// LS Electric XG5000 project: 555
// PLC LSPLC

PROGRAM E2E_PICKNPLACE (task: 스캔 프로그램)

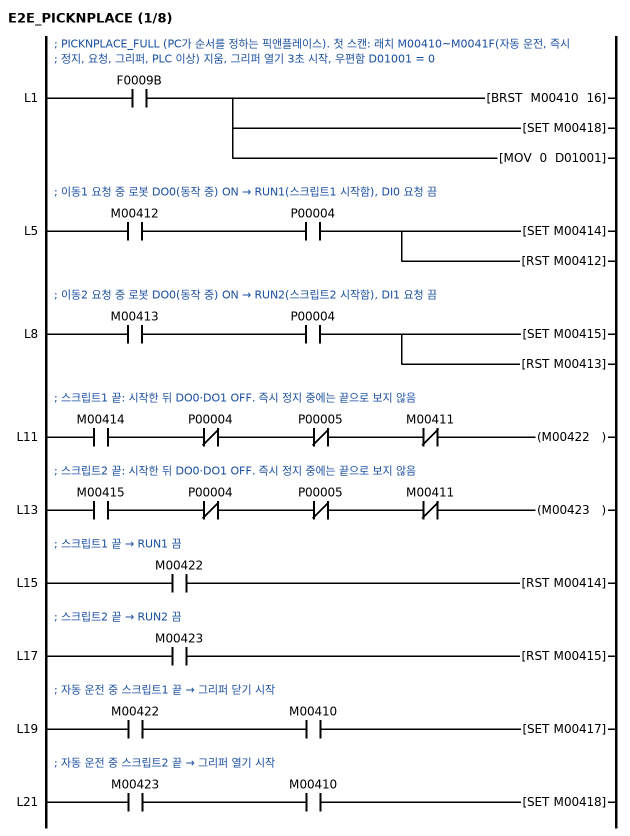
// PICKNPLACE_FULL (PC가 순서를 정하는 픽앤플레이스). 첫 스캔: 래치 M00410~M0041F(자동 운전, 즉시 정지, 요청, 그리퍼, PLC 이상) 지움, 그리퍼 열기 3초 시작, 우편함 D01001 = 0
; L1
LOAD      F0009B
BRST      M00410 16
SET       M00418
MOV       0 D01001
// 이동1 요청 중 로봇 DO0(동작 중) ON → RUN1(스크립트1 시작함), DI0 요청 끔
; L5
LOAD      M00412
AND       P00004
SET       M00414
RST       M00412
// 이동2 요청 중 로봇 DO0(동작 중) ON → RUN2(스크립트2 시작함), DI1 요청 끔
; L8
LOAD      M00413
AND       P00004
SET       M00415
RST       M00413
// 스크립트1 끝: 시작한 뒤 DO0·DO1 OFF. 즉시 정지 중에는 끝으로 보지 않음
; L11
LOAD      M00414
AND NOT   P00004
AND NOT   P00005
AND NOT   M00411
OUT       M00422
// 스크립트2 끝: 시작한 뒤 DO0·DO1 OFF. 즉시 정지 중에는 끝으로 보지 않음
; L13
LOAD      M00415
AND NOT   P00004
AND NOT   P00005
AND NOT   M00411
OUT       M00423
// 스크립트1 끝 → RUN1 끔
; L15
LOAD      M00422
RST       M00414
// 스크립트2 끝 → RUN2 끔
; L17
LOAD      M00423
RST       M00415
// 자동 운전 중 스크립트1 끝 → 그리퍼 닫기 시작
; L19
LOAD      M00422
AND       M00410
SET       M00417
// 자동 운전 중 스크립트2 끝 → 그리퍼 열기 시작
; L21
LOAD      M00423
AND       M00410
SET       M00418

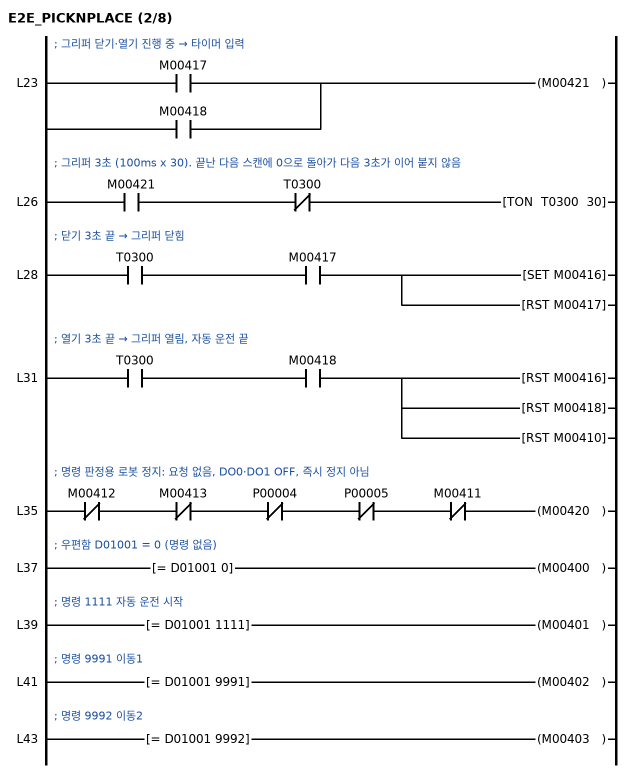
// 그리퍼 닫기·열기 진행 중 → 타이머 입력
; L23
LOAD      M00417
OR        M00418
OUT       M00421
// 그리퍼 3초 (100ms x 30). 끝난 다음 스캔에 0으로 돌아가 다음 3초가 이어 붙지 않음
; L26
LOAD      M00421
AND NOT   T0300
TON       T0300 30
// 닫기 3초 끝 → 그리퍼 닫힘
; L28
LOAD      T0300
AND       M00417
SET       M00416
RST       M00417
// 열기 3초 끝 → 그리퍼 열림, 자동 운전 끝
; L31
LOAD      T0300
AND       M00418
RST       M00416
RST       M00418
RST       M00410
// 명령 판정용 로봇 정지: 요청 없음, DO0·DO1 OFF, 즉시 정지 아님
; L35
LOAD NOT  M00412
AND NOT   M00413
AND NOT   P00004
AND NOT   P00005
AND NOT   M00411
OUT       M00420
// 우편함 D01001 = 0 (명령 없음)
; L37
LOAD=     D01001 0
OUT       M00400
// 명령 1111 자동 운전 시작
; L39
LOAD=     D01001 1111
OUT       M00401
// 명령 9991 이동1
; L41
LOAD=     D01001 9991
OUT       M00402
// 명령 9992 이동2
; L43
LOAD=     D01001 9992
OUT       M00403

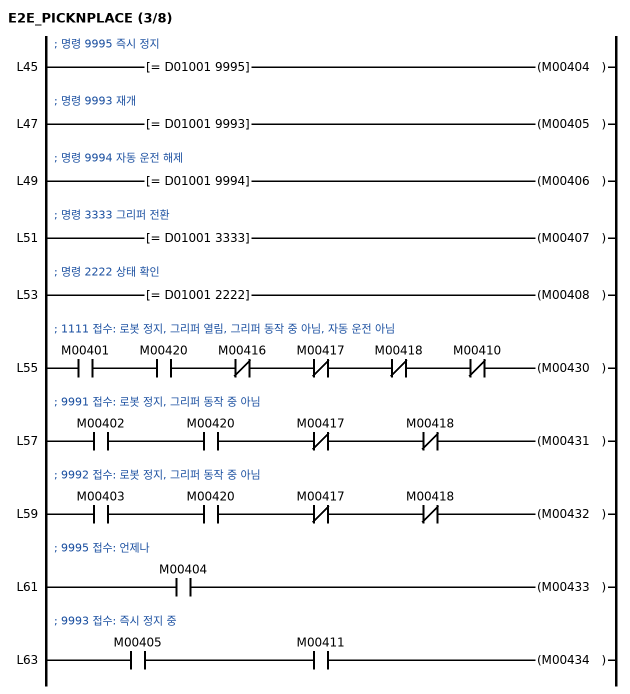
// 명령 9995 즉시 정지
; L45
LOAD=     D01001 9995
OUT       M00404
// 명령 9993 재개
; L47
LOAD=     D01001 9993
OUT       M00405
// 명령 9994 자동 운전 해제
; L49
LOAD=     D01001 9994
OUT       M00406
// 명령 3333 그리퍼 전환
; L51
LOAD=     D01001 3333
OUT       M00407
// 명령 2222 상태 확인
; L53
LOAD=     D01001 2222
OUT       M00408
// 1111 접수: 로봇 정지, 그리퍼 열림, 그리퍼 동작 중 아님, 자동 운전 아님
; L55
LOAD      M00401
AND       M00420
AND NOT   M00416
AND NOT   M00417
AND NOT   M00418
AND NOT   M00410
OUT       M00430
// 9991 접수: 로봇 정지, 그리퍼 동작 중 아님
; L57
LOAD      M00402
AND       M00420
AND NOT   M00417
AND NOT   M00418
OUT       M00431
// 9992 접수: 로봇 정지, 그리퍼 동작 중 아님
; L59
LOAD      M00403
AND       M00420
AND NOT   M00417
AND NOT   M00418
OUT       M00432
// 9995 접수: 언제나
; L61
LOAD      M00404
OUT       M00433
// 9993 접수: 즉시 정지 중
; L63
LOAD      M00405
AND       M00411
OUT       M00434

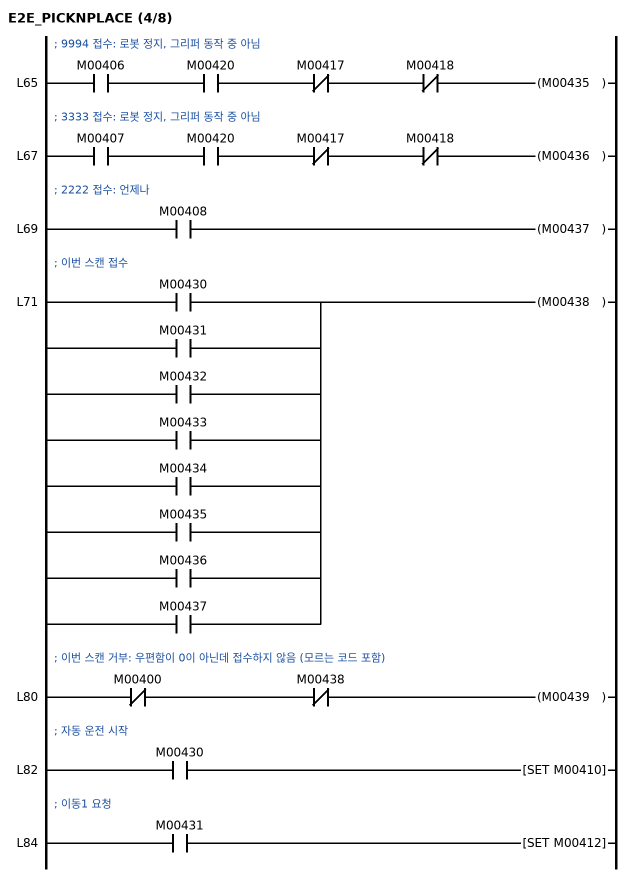
// 9994 접수: 로봇 정지, 그리퍼 동작 중 아님
; L65
LOAD      M00406
AND       M00420
AND NOT   M00417
AND NOT   M00418
OUT       M00435
// 3333 접수: 로봇 정지, 그리퍼 동작 중 아님
; L67
LOAD      M00407
AND       M00420
AND NOT   M00417
AND NOT   M00418
OUT       M00436
// 2222 접수: 언제나
; L69
LOAD      M00408
OUT       M00437
// 이번 스캔 접수
; L71
LOAD      M00430
OR        M00431
OR        M00432
OR        M00433
OR        M00434
OR        M00435
OR        M00436
OR        M00437
OUT       M00438
// 이번 스캔 거부: 우편함이 0이 아닌데 접수하지 않음 (모르는 코드 포함)
; L80
LOAD NOT  M00400
AND NOT   M00438
OUT       M00439
// 자동 운전 시작
; L82
LOAD      M00430
SET       M00410
// 이동1 요청
; L84
LOAD      M00431
SET       M00412

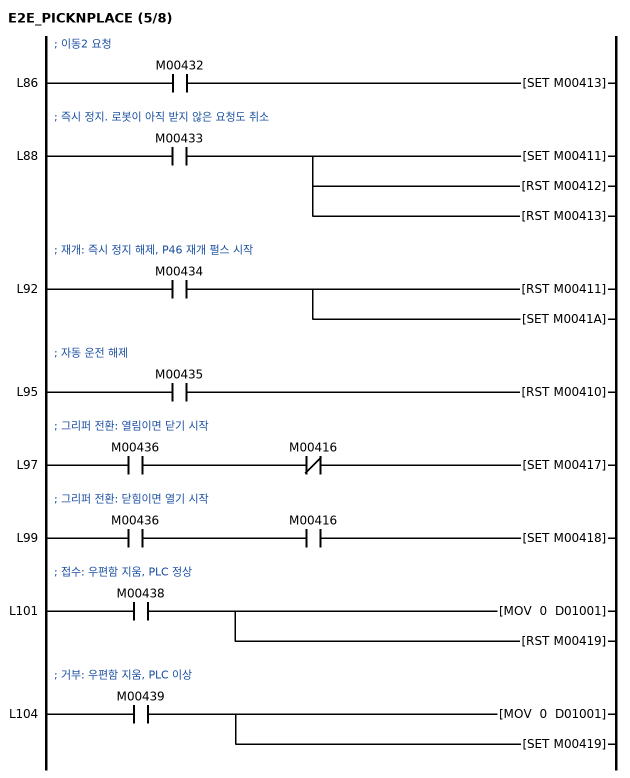
// 이동2 요청
; L86
LOAD      M00432
SET       M00413
// 즉시 정지. 로봇이 아직 받지 않은 요청도 취소
; L88
LOAD      M00433
SET       M00411
RST       M00412
RST       M00413
// 재개: 즉시 정지 해제, P46 재개 펄스 시작
; L92
LOAD      M00434
RST       M00411
SET       M0041A
// 자동 운전 해제
; L95
LOAD      M00435
RST       M00410
// 그리퍼 전환: 열림이면 닫기 시작
; L97
LOAD      M00436
AND NOT   M00416
SET       M00417
// 그리퍼 전환: 닫힘이면 열기 시작
; L99
LOAD      M00436
AND       M00416
SET       M00418
// 접수: 우편함 지움, PLC 정상
; L101
LOAD      M00438
MOV       0 D01001
RST       M00419
// 거부: 우편함 지움, PLC 이상
; L104
LOAD      M00439
MOV       0 D01001
SET       M00419

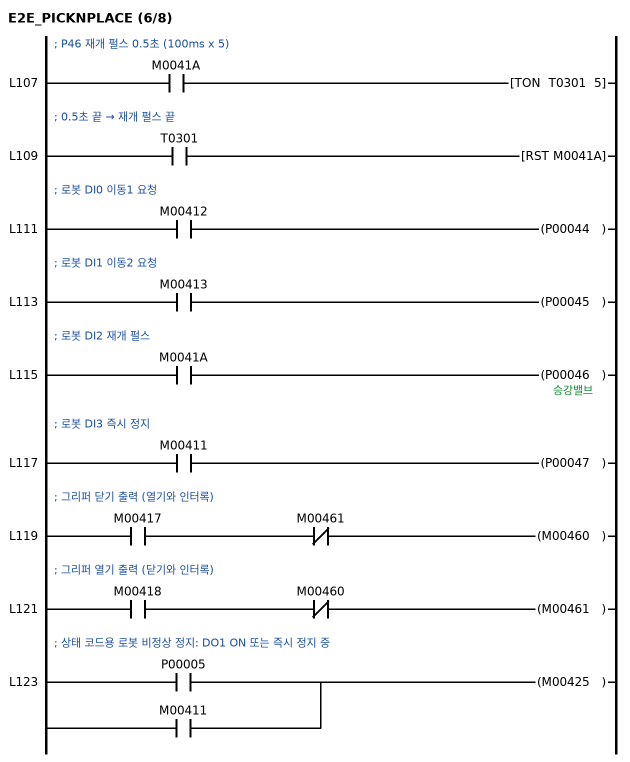
// P46 재개 펄스 0.5초 (100ms x 5)
; L107
LOAD      M0041A
TON       T0301 5
// 0.5초 끝 → 재개 펄스 끝
; L109
LOAD      T0301
RST       M0041A
// 로봇 DI0 이동1 요청
; L111
LOAD      M00412
OUT       P00044
// 로봇 DI1 이동2 요청
; L113
LOAD      M00413
OUT       P00045
// 로봇 DI2 재개 펄스
; L115
LOAD      M0041A
OUT       P00046	// 승강밸브
// 로봇 DI3 즉시 정지
; L117
LOAD      M00411
OUT       P00047
// 그리퍼 닫기 출력 (열기와 인터록)
; L119
LOAD      M00417
AND NOT   M00461
OUT       M00460
// 그리퍼 열기 출력 (닫기와 인터록)
; L121
LOAD      M00418
AND NOT   M00460
OUT       M00461
// 상태 코드용 로봇 비정상 정지: DO1 ON 또는 즉시 정지 중
; L123
LOAD      P00005
OR        M00411
OUT       M00425

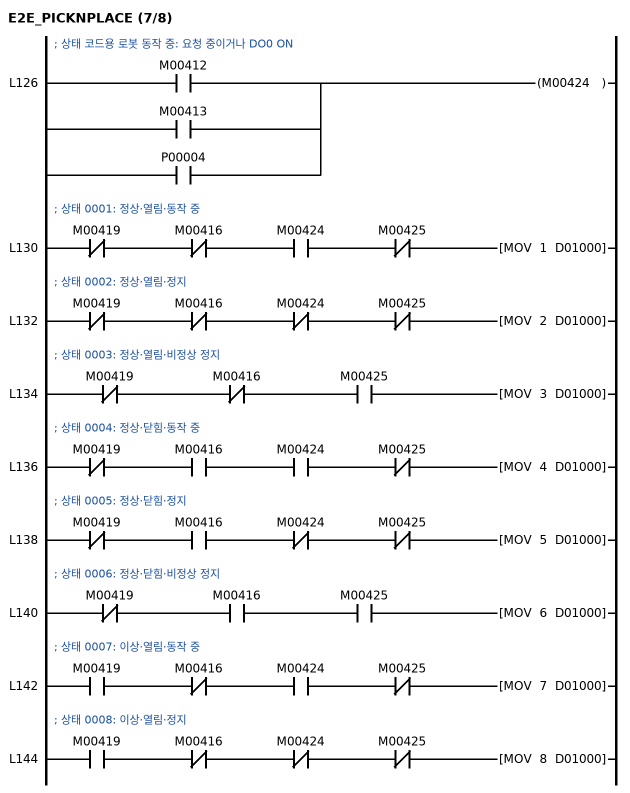
// 상태 코드용 로봇 동작 중: 요청 중이거나 DO0 ON
; L126
LOAD      M00412
OR        M00413
OR        P00004
OUT       M00424
// 상태 0001: 정상·열림·동작 중
; L130
LOAD NOT  M00419
AND NOT   M00416
AND       M00424
AND NOT   M00425
MOV       1 D01000
// 상태 0002: 정상·열림·정지
; L132
LOAD NOT  M00419
AND NOT   M00416
AND NOT   M00424
AND NOT   M00425
MOV       2 D01000
// 상태 0003: 정상·열림·비정상 정지
; L134
LOAD NOT  M00419
AND NOT   M00416
AND       M00425
MOV       3 D01000
// 상태 0004: 정상·닫힘·동작 중
; L136
LOAD NOT  M00419
AND       M00416
AND       M00424
AND NOT   M00425
MOV       4 D01000
// 상태 0005: 정상·닫힘·정지
; L138
LOAD NOT  M00419
AND       M00416
AND NOT   M00424
AND NOT   M00425
MOV       5 D01000
// 상태 0006: 정상·닫힘·비정상 정지
; L140
LOAD NOT  M00419
AND       M00416
AND       M00425
MOV       6 D01000
// 상태 0007: 이상·열림·동작 중
; L142
LOAD      M00419
AND NOT   M00416
AND       M00424
AND NOT   M00425
MOV       7 D01000
// 상태 0008: 이상·열림·정지
; L144
LOAD      M00419
AND NOT   M00416
AND NOT   M00424
AND NOT   M00425
MOV       8 D01000

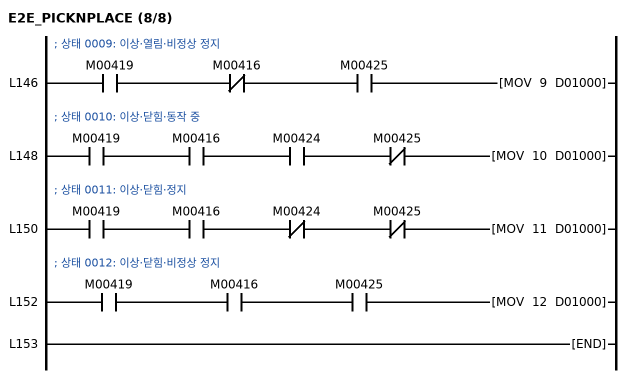
// 상태 0009: 이상·열림·비정상 정지
; L146
LOAD      M00419
AND NOT   M00416
AND       M00425
MOV       9 D01000
// 상태 0010: 이상·닫힘·동작 중
; L148
LOAD      M00419
AND       M00416
AND       M00424
AND NOT   M00425
MOV       10 D01000
// 상태 0011: 이상·닫힘·정지
; L150
LOAD      M00419
AND       M00416
AND NOT   M00424
AND NOT   M00425
MOV       11 D01000
// 상태 0012: 이상·닫힘·비정상 정지
; L152
LOAD      M00419
AND       M00416
AND       M00425
MOV       12 D01000
; L153
END

VARIABLES AND COMMENTS (devices not used above)
P00041	BIT	GL1
P00000	BIT	PB1
P00001	BIT	PB2
P00042	BIT	YL1
M00103	BIT	상승1
P00007	BIT	상승단
M00100	BIT	원점대기
M00102	BIT	잡기대기
T0100	BIT/WORD	타이머_1초
M00101	BIT	하강1
P00008	BIT	하강단